// TIA Portal V20 export
// export: Created 2026-10-11T05:32:37.6267366Z, ExportSetting WithDefaults, DisplayName Totally Integrated Automation Portal, DisplayVersion V20, DisplayName TIA Portal Openness, DisplayVersion V20, DisplayName TIA Portal Teamcenter Gateway, DisplayVersion V20, DisplayName TIA Portal Version Control Interface, DisplayVersion V20, DisplayName SINAMICS Startdrive Advanced, DisplayVersion V20 SP1 Update 2, DisplayName SINAMICS Startdrive G110M, G120, G120C, G120D, G120P, G115D, DisplayVersion V20 SP1 Update 2, DisplayName SINAMICS Startdrive G130, G150, S120, S150, SINAMICS MV, G220, S200, S210, DisplayVersion V20 SP1 Update 2, DisplayName STEP 7 Professional, DisplayVersion V20, DisplayName STEP 7 Safety, DisplayVersion V20, DisplayName WinCC Basic/Comfort/Advanced, DisplayVersion V20, DisplayName WinCC Professional, DisplayVersion V20, DisplayName WinCC Unified, DisplayVersion V20
FUNCTION "FRK_PartAborted" : Void   // FC41, SCL
{ S7_Optimized_Access := 'TRUE' }
VERSION : 0.1
// stored: AutoNumber true, IsIECCheckEnabled false, SetENOAutomatically false, UDAEnableTagReadback false
   VAR_IN_OUT
      Core : "FRK_Core";
      Unit : "FRK_Unit";
      Status : "ST_ModuleStatus";
      Part : "ST_PartContext";
      History : Array[1..16] of "ST_Diagnostic";
      Head : Int;
   END_VAR
BEGIN

   IF #Unit.CarrierIndex = 0 OR NOT #Part.Present THEN
       RETURN;
   END_IF;
   #Part.Result.Verdict := 0;
   IF #Core.Exec = 3 AND #Part.Result.ReasonCode = 0 THEN
       #Part.Result.ReasonCode := #Status.Diagnostic.ReasonCode;
   END_IF;
   "FRK_PartEvent"(History := #History,
                   Head := #Head,
                   Reason := 2027,
                   Uid := #Part.Uid,
                   SourcePath := #Status.Name);
   #Part.Present := FALSE;
END_FUNCTION
